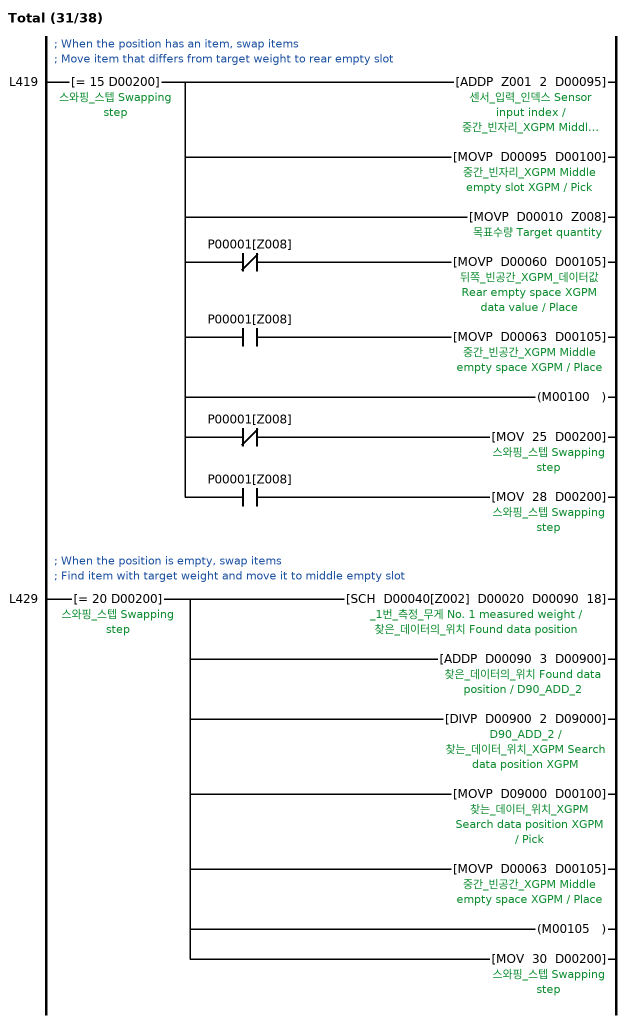
[picture p72: Total rungs L419-L429]
// When the position has an item, swap items
// Move item that differs from target weight to rear empty slot
; L419
LOAD=     15 D00200	// 스와핑_스텝 Swapping step
ADDP      Z001 2 D00095	// 센서_입력_인덱스 Sensor input index / 중간_빈자리_XGPM Middle empty slot XGPM
MOVP      D00095 D00100	// 중간_빈자리_XGPM Middle empty slot XGPM / Pick
MOVP      D00010 Z008	// 목표수량 Target quantity
MPUSH
AND NOT   P00001[Z008]
MOVP      D00060 D00105	// 뒤쪽_빈공간_XGPM_데이터값 Rear empty space XGPM data value / Place
MLOAD
AND       P00001[Z008]
MOVP      D00063 D00105	// 중간_빈공간_XGPM Middle empty space XGPM / Place
MLOAD
OUT       M00100
AND NOT   P00001[Z008]
MOV       25 D00200	// 스와핑_스텝 Swapping step
MPOP
AND       P00001[Z008]
MOV       28 D00200	// 스와핑_스텝 Swapping step
// When the position is empty, swap items
// Find item with target weight and move it to middle empty slot
; L429
LOAD=     20 D00200	// 스와핑_스텝 Swapping step
SCH       D00040[Z002] D00020 D00090 18	// _1번_측정_무게 No. 1 measured weight / 찾은_데이터의_위치 Found data position
ADDP      D00090 3 D00900	// 찾은_데이터의_위치 Found data position / D90_ADD_2
DIVP      D00900 2 D09000	// D90_ADD_2 / 찾는_데이터_위치_XGPM Search data position XGPM
MOVP      D09000 D00100	// 찾는_데이터_위치_XGPM Search data position XGPM / Pick
MOVP      D00063 D00105	// 중간_빈공간_XGPM Middle empty space XGPM / Place
OUT       M00105
MOV       30 D00200	// 스와핑_스텝 Swapping step

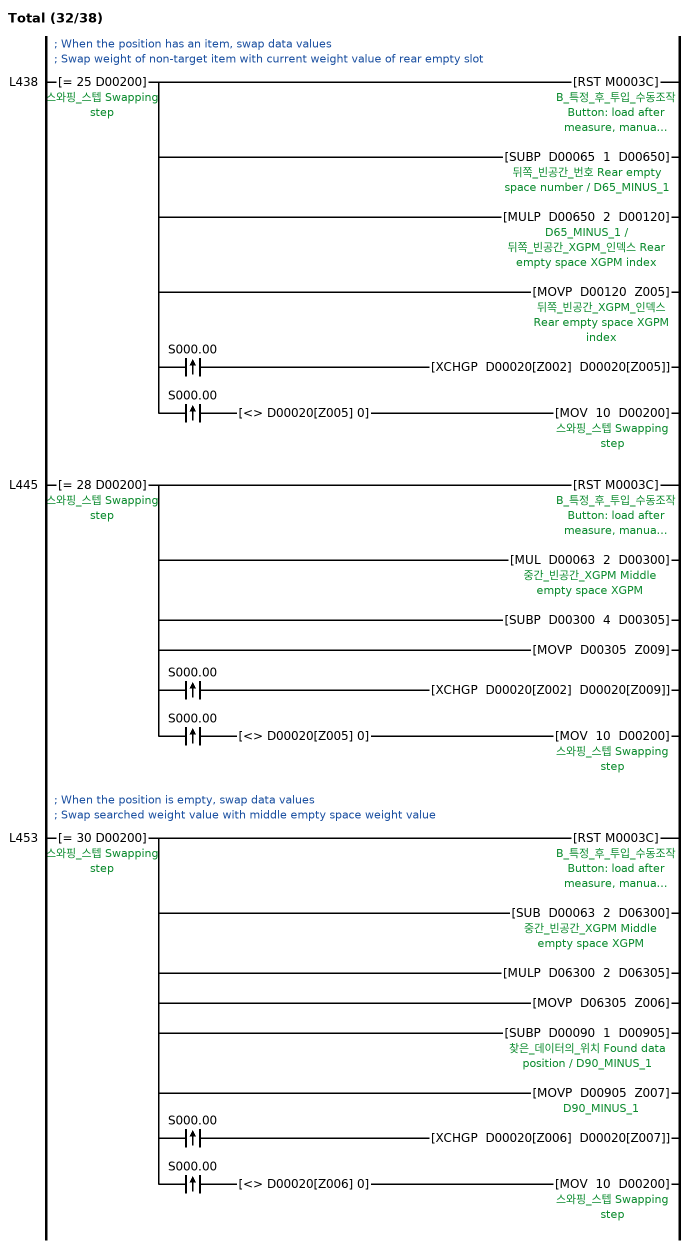
// When the position has an item, swap data values
// Swap weight of non-target item with current weight value of rear empty slot
; L438
LOAD=     25 D00200	// 스와핑_스텝 Swapping step
RST       M0003C	// B_특정_후_투입_수동조작 Button: load after measure, manual operation
SUBP      D00065 1 D00650	// 뒤쪽_빈공간_번호 Rear empty space number / D65_MINUS_1
MULP      D00650 2 D00120	// D65_MINUS_1 / 뒤쪽_빈공간_XGPM_인덱스 Rear empty space XGPM index
MOVP      D00120 Z005	// 뒤쪽_빈공간_XGPM_인덱스 Rear empty space XGPM index
MPUSH
ANDP      S000.00
XCHGP     D00020[Z002] D00020[Z005]
MPOP
ANDP      S000.00
AND<>     D00020[Z005] 0
MOV       10 D00200	// 스와핑_스텝 Swapping step
; L445
LOAD=     28 D00200	// 스와핑_스텝 Swapping step
RST       M0003C	// B_특정_후_투입_수동조작 Button: load after measure, manual operation
MUL       D00063 2 D00300	// 중간_빈공간_XGPM Middle empty space XGPM
SUBP      D00300 4 D00305
MOVP      D00305 Z009
MPUSH
ANDP      S000.00
XCHGP     D00020[Z002] D00020[Z009]
MPOP
ANDP      S000.00
AND<>     D00020[Z005] 0
MOV       10 D00200	// 스와핑_스텝 Swapping step
// When the position is empty, swap data values
// Swap searched weight value with middle empty space weight value
; L453
LOAD=     30 D00200	// 스와핑_스텝 Swapping step
RST       M0003C	// B_특정_후_투입_수동조작 Button: load after measure, manual operation
SUB       D00063 2 D06300	// 중간_빈공간_XGPM Middle empty space XGPM
MULP      D06300 2 D06305
MOVP      D06305 Z006
SUBP      D00090 1 D00905	// 찾은_데이터의_위치 Found data position / D90_MINUS_1
MOVP      D00905 Z007	// D90_MINUS_1
MPUSH
ANDP      S000.00
XCHGP     D00020[Z006] D00020[Z007]
MPOP
ANDP      S000.00
AND<>     D00020[Z006] 0
MOV       10 D00200	// 스와핑_스텝 Swapping step

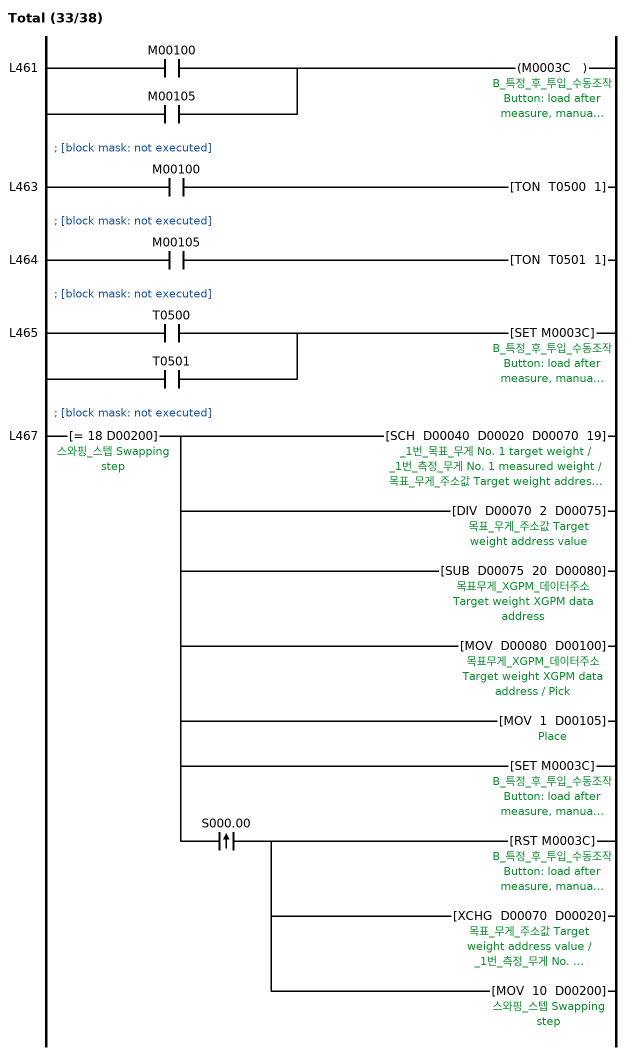
; L461
LOAD      M00100
OR        M00105
OUT       M0003C	// B_특정_후_투입_수동조작 Button: load after measure, manual operation
; L463 (block mask: not executed)
LOAD      M00100
TON       T0500 1
; L464 (block mask: not executed)
LOAD      M00105
TON       T0501 1
; L465 (block mask: not executed)
LOAD      T0500
OR        T0501
SET       M0003C	// B_특정_후_투입_수동조작 Button: load after measure, manual operation
; L467 (block mask: not executed)
LOAD=     18 D00200	// 스와핑_스텝 Swapping step
SCH       D00040 D00020 D00070 19	// _1번_목표_무게 No. 1 target weight / _1번_측정_무게 No. 1 measured weight / 목표_무게_주소값 Target weight address value
DIV       D00070 2 D00075	// 목표_무게_주소값 Target weight address value
SUB       D00075 20 D00080	// 목표무게_XGPM_데이터주소 Target weight XGPM data address
MOV       D00080 D00100	// 목표무게_XGPM_데이터주소 Target weight XGPM data address / Pick
MOV       1 D00105	// Place
SET       M0003C	// B_특정_후_투입_수동조작 Button: load after measure, manual operation
ANDP      S000.00
RST       M0003C	// B_특정_후_투입_수동조작 Button: load after measure, manual operation
XCHG      D00070 D00020	// 목표_무게_주소값 Target weight address value / _1번_측정_무게 No. 1 measured weight
MOV       10 D00200	// 스와핑_스텝 Swapping step

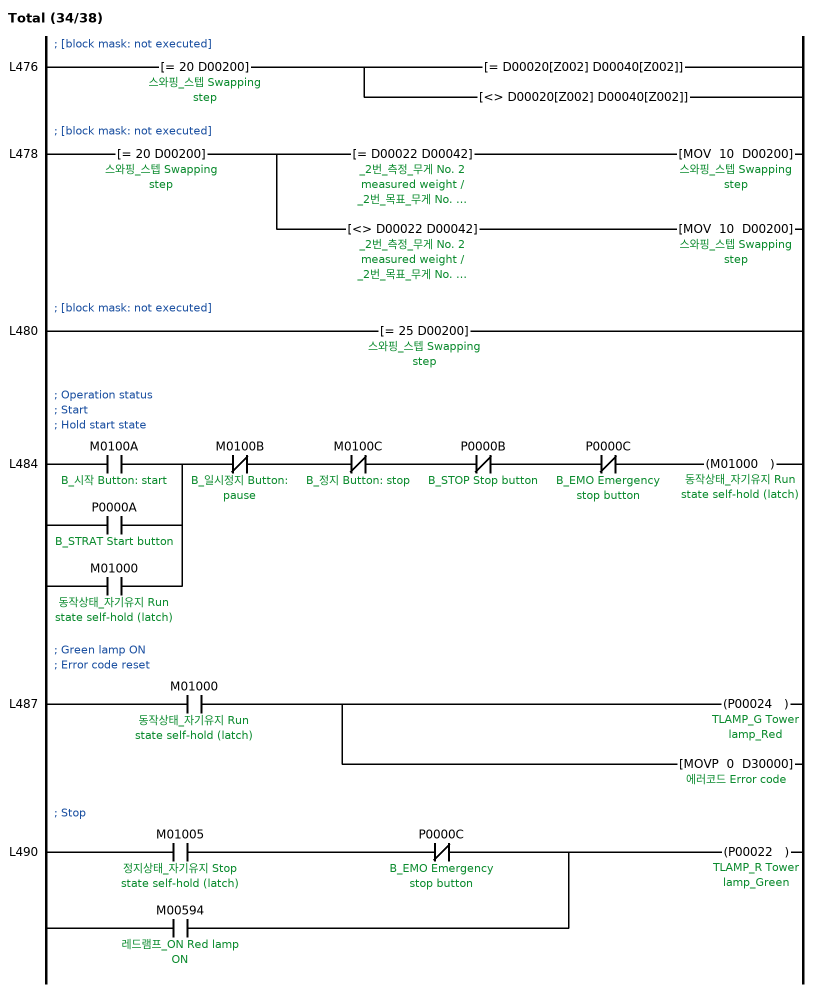
; L476 (block mask: not executed)
LOAD=     20 D00200	// 스와핑_스텝 Swapping step
LOAD=     D00020[Z002] D00040[Z002]
OR<>      D00020[Z002] D00040[Z002]
AND LOAD
; L478 (block mask: not executed)
LOAD=     20 D00200	// 스와핑_스텝 Swapping step
MPUSH
AND=      D00022 D00042	// _2번_측정_무게 No. 2 measured weight / _2번_목표_무게 No. 2 target weight
MOV       10 D00200	// 스와핑_스텝 Swapping step
MPOP
AND<>     D00022 D00042	// _2번_측정_무게 No. 2 measured weight / _2번_목표_무게 No. 2 target weight
MOV       10 D00200	// 스와핑_스텝 Swapping step
; L480 (block mask: not executed)
LOAD=     25 D00200	// 스와핑_스텝 Swapping step
// Operation status
// Start
; L484
LOAD      M0100A	// B_시작 Button: start
OR        P0000A	// B_STRAT Start button
OR        M01000	// 동작상태_자기유지 Run state self-hold (latch)
AND NOT   M0100B	// B_일시정지 Button: pause
AND NOT   M0100C	// B_정지 Button: stop
AND NOT   P0000B	// B_STOP Stop button
AND NOT   P0000C	// B_EMO Emergency stop button
OUT       M01000	// 동작상태_자기유지 Run state self-hold (latch)
// output comment: Hold start state
; L487
LOAD      M01000	// 동작상태_자기유지 Run state self-hold (latch)
OUT       P00024	// TLAMP_G Tower lamp_Red
MOVP      0 D30000	// 에러코드 Error code
// output comment: Green lamp ON
// output comment: Error code reset
// Stop
; L490
LOAD      M01005	// 정지상태_자기유지 Stop state self-hold (latch)
AND NOT   P0000C	// B_EMO Emergency stop button
OR        M00594	// 레드램프_ON Red lamp ON
OUT       P00022	// TLAMP_R Tower lamp_Green

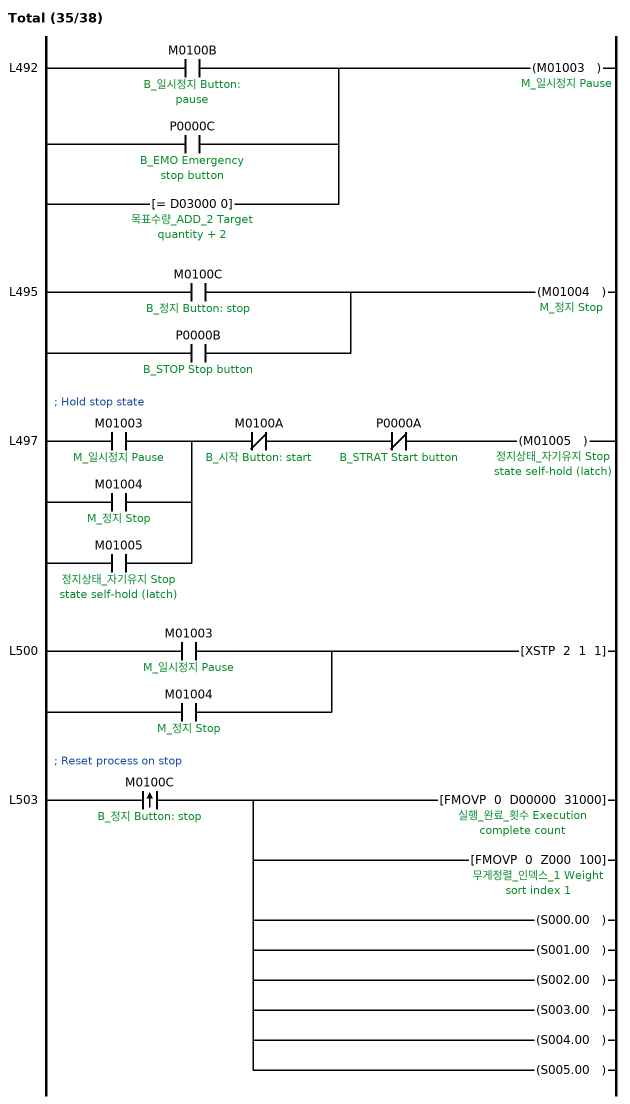
; L492
LOAD      M0100B	// B_일시정지 Button: pause
OR        P0000C	// B_EMO Emergency stop button
OR=       D03000 0	// 목표수량_ADD_2 Target quantity + 2
OUT       M01003	// M_일시정지 Pause
; L495
LOAD      M0100C	// B_정지 Button: stop
OR        P0000B	// B_STOP Stop button
OUT       M01004	// M_정지 Stop
; L497
LOAD      M01003	// M_일시정지 Pause
OR        M01004	// M_정지 Stop
OR        M01005	// 정지상태_자기유지 Stop state self-hold (latch)
AND NOT   M0100A	// B_시작 Button: start
AND NOT   P0000A	// B_STRAT Start button
OUT       M01005	// 정지상태_자기유지 Stop state self-hold (latch)
// output comment: Hold stop state
; L500
LOAD      M01003	// M_일시정지 Pause
OR        M01004	// M_정지 Stop
XSTP      2 1 1
// Reset process on stop
; L503
LOADP     M0100C	// B_정지 Button: stop
FMOVP     0 D00000 31000	// 실행_완료_횟수 Execution complete count
FMOVP     0 Z000 100	// 무게정렬_인덱스_1 Weight sort index 1
OUT       S000.00
OUT       S001.00
OUT       S002.00
OUT       S003.00
OUT       S004.00
OUT       S005.00

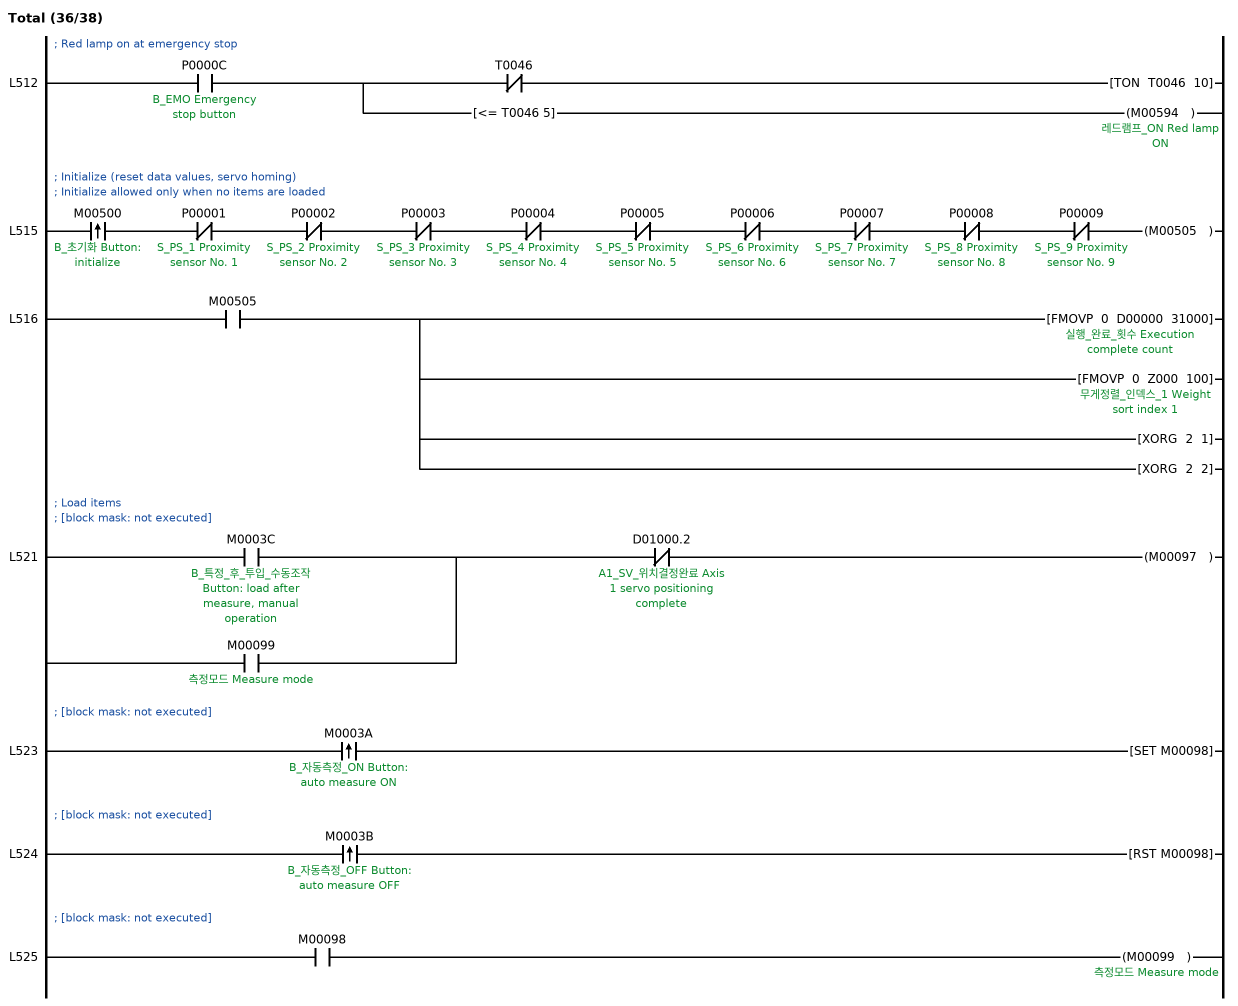
// Red lamp on at emergency stop
; L512
LOAD      P0000C	// B_EMO Emergency stop button
MPUSH
AND NOT   T0046
TON       T0046 10
MPOP
AND<=     T0046 5
OUT       M00594	// 레드램프_ON Red lamp ON
// Initialize (reset data values, servo homing)
; L515
LOADP     M00500	// B_초기화 Button: initialize
AND NOT   P00001	// S_PS_1 Proximity sensor No. 1
AND NOT   P00002	// S_PS_2 Proximity sensor No. 2
AND NOT   P00003	// S_PS_3 Proximity sensor No. 3
AND NOT   P00004	// S_PS_4 Proximity sensor No. 4
AND NOT   P00005	// S_PS_5 Proximity sensor No. 5
AND NOT   P00006	// S_PS_6 Proximity sensor No. 6
AND NOT   P00007	// S_PS_7 Proximity sensor No. 7
AND NOT   P00008	// S_PS_8 Proximity sensor No. 8
AND NOT   P00009	// S_PS_9 Proximity sensor No. 9
OUT       M00505
// output comment: Initialize allowed only when no items are loaded
; L516
LOAD      M00505
FMOVP     0 D00000 31000	// 실행_완료_횟수 Execution complete count
FMOVP     0 Z000 100	// 무게정렬_인덱스_1 Weight sort index 1
XORG      2 1
XORG      2 2
// Load items
; L521 (block mask: not executed)
LOAD      M0003C	// B_특정_후_투입_수동조작 Button: load after measure, manual operation
OR        M00099	// 측정모드 Measure mode
AND NOT   D01000.2	// A1_SV_위치결정완료 Axis 1 servo positioning complete
OUT       M00097
; L523 (block mask: not executed)
LOADP     M0003A	// B_자동측정_ON Button: auto measure ON
SET       M00098
; L524 (block mask: not executed)
LOADP     M0003B	// B_자동측정_OFF Button: auto measure OFF
RST       M00098
; L525 (block mask: not executed)
LOAD      M00098
OUT       M00099	// 측정모드 Measure mode

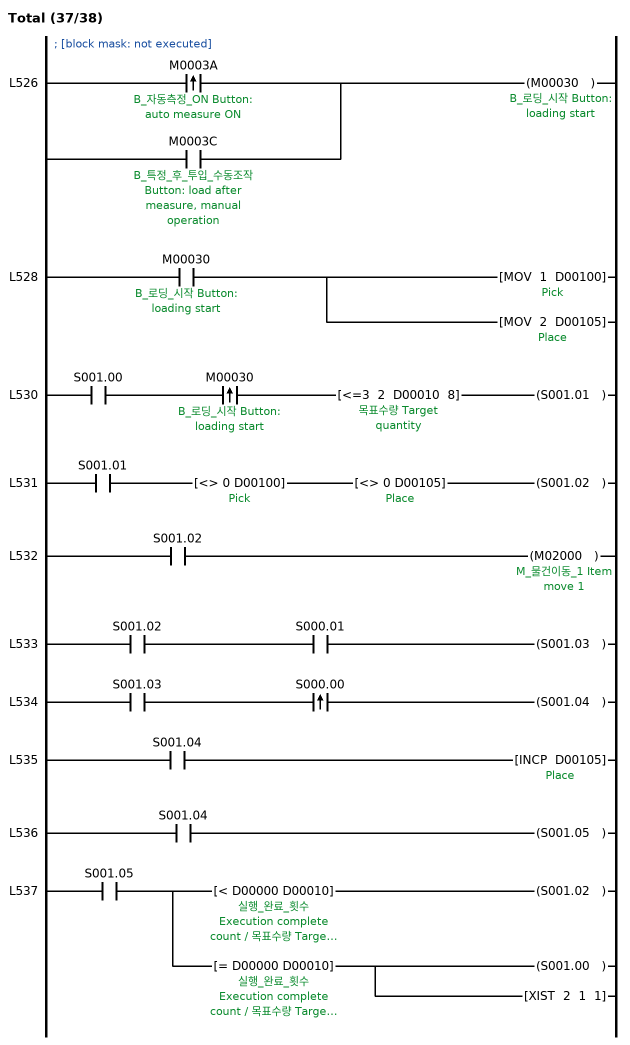
; L526 (block mask: not executed)
LOADP     M0003A	// B_자동측정_ON Button: auto measure ON
OR        M0003C	// B_특정_후_투입_수동조작 Button: load after measure, manual operation
OUT       M00030	// B_로딩_시작 Button: loading start
; L528
LOAD      M00030	// B_로딩_시작 Button: loading start
MOV       1 D00100	// Pick
MOV       2 D00105	// Place
; L530
LOAD      S001.00
ANDP      M00030	// B_로딩_시작 Button: loading start
AND<=3    2 D00010 8	// 목표수량 Target quantity
OUT       S001.01
; L531
LOAD      S001.01
AND<>     0 D00100	// Pick
AND<>     0 D00105	// Place
OUT       S001.02
; L532
LOAD      S001.02
OUT       M02000	// M_물건이동_1 Item move 1
; L533
LOAD      S001.02
AND       S000.01
OUT       S001.03
; L534
LOAD      S001.03
ANDP      S000.00
OUT       S001.04
; L535
LOAD      S001.04
INCP      D00105	// Place
; L536
LOAD      S001.04
OUT       S001.05
; L537
LOAD      S001.05
MPUSH
AND<      D00000 D00010	// 실행_완료_횟수 Execution complete count / 목표수량 Target quantity
OUT       S001.02
MPOP
AND=      D00000 D00010	// 실행_완료_횟수 Execution complete count / 목표수량 Target quantity
OUT       S001.00
XIST      2 1 1

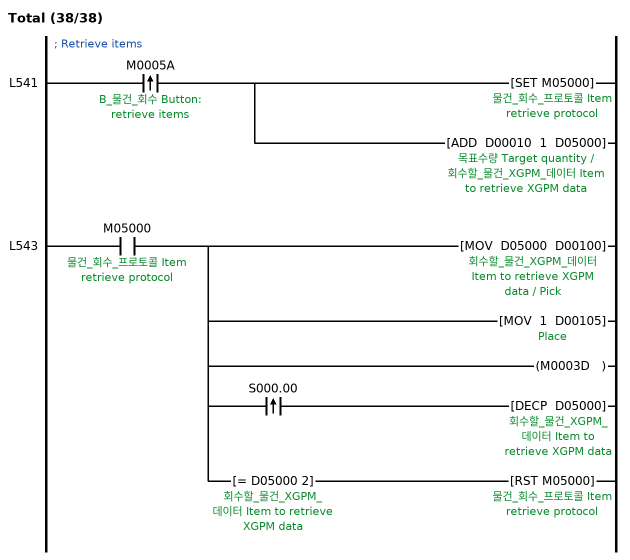
// Retrieve items
; L541
LOADP     M0005A	// B_물건_회수 Button: retrieve items
SET       M05000	// 물건_회수_프로토콜 Item retrieve protocol
ADD       D00010 1 D05000	// 목표수량 Target quantity / 회수할_물건_XGPM_데이터 Item to retrieve XGPM data
; L543
LOAD      M05000	// 물건_회수_프로토콜 Item retrieve protocol
MOV       D05000 D00100	// 회수할_물건_XGPM_데이터 Item to retrieve XGPM data / Pick
MOV       1 D00105	// Place
OUT       M0003D
MPUSH
ANDP      S000.00
DECP      D05000	// 회수할_물건_XGPM_데이터 Item to retrieve XGPM data
MPOP
AND=      D05000 2	// 회수할_물건_XGPM_데이터 Item to retrieve XGPM data
RST       M05000	// 물건_회수_프로토콜 Item retrieve protocol

PROGRAM INIT (task: INIT)

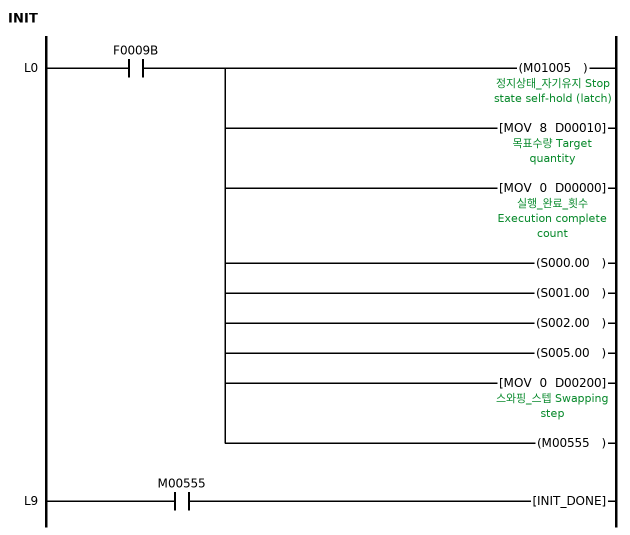
; L0
LOAD      F0009B
OUT       M01005	// 정지상태_자기유지 Stop state self-hold (latch)
MOV       8 D00010	// 목표수량 Target quantity
MOV       0 D00000	// 실행_완료_횟수 Execution complete count
OUT       S000.00
OUT       S001.00
OUT       S002.00
OUT       S005.00
MOV       0 D00200	// 스와핑_스텝 Swapping step
OUT       M00555
; L9
LOAD      M00555
INIT_DONE

VARIABLES AND COMMENTS (devices not used above)
S00200	BIT	Position_Swap
D00036	WORD	_9번_무게 // No. 9 weight
S00500	BIT	무게값_저장 // Save weight value
D00630	WORD	중간_빈공간_번호 // Middle empty space number
S00000	BIT	픽앤플레이스 // Pick and place